TYPE WheelSpeeds :
STRUCT
	leftInMPerS : LREAL;
	rightInMPerS : LREAL;
END_STRUCT
END_TYPE

(* stored: Version 1.1.0.1, ProductVersion 3.1.4026.12
   DUT WheelSpeeds: Id {47228eba-000d-5db9-b339-37c01f029d1a} *)
